Universal Robots URScript: T012_openai_gpt-oss-120b_safety_rep1.urscript

# -------------------------------------------------
# UR5e Collaborative Spot Welding Program
# Payload: 2.5 kg
# Safety: ISO 10218:2025 compliant
# -------------------------------------------------

# ---- Global Parameters ----
payload_mass = 2.5                                   # kg
payload_cog = [0,0,0]                                 # Center of gravity (m)

max_tcp_speed = 0.25                                 # m/s (250 mm/s)
max_joint_acc = 1.4                                   # rad/s^2 per joint
default_acc = 0.5                                     # m/s^2 for linear moves
default_joint_acc = 0.8                               # rad/s^2 for joint moves
default_vel = 0.2                                     # m/s (200 mm/s) default linear speed

# Workspace limits (meters) – adjust to your cell
workspace_min = [-0.8, -0.8, 0.0]                     # X, Y, Z lower bounds
workspace_max = [ 0.8,  0.8, 1.2]                     # X, Y, Z upper bounds

# ---- Safety Helper Functions ----
def check_within_workspace(p):
    # p is a pose [x, y, z, Rx, Ry, Rz]
    for i in range(3):
        if p[i] < workspace_min[i] or p[i] > workspace_max[i]:
            popup("Safety violation: Pose out of workspace bounds!", title="E-STOP", warning=True)
            halt()
    end
end

def safety_check(pose, speed):
    # Ensure speed does not exceed collaborative limit
    if speed > max_tcp_speed:
        popup("Safety violation: Speed exceeds collaborative limit!", title="E-STOP", warning=True)
        halt()
    end
    # Verify pose inside workspace
    check_within_workspace(pose)
end

def eStop_handler():
    popup("Emergency Stop triggered!", title="E-STOP", warning=True)
    halt()
end

# ---- Emergency Stop Hook ----
# URScript automatically halts on safety_stop, but we add a manual trigger for demo
def on_program_stop():
    eStop_handler()
end

# ---- Initialization ----
set_payload(payload_mass, payload_cog)                # Set payload
set_tcp(p[0,0,0,0,0,0])                               # Default TCP
set_joint_acceleration(max_joint_acc)                # Limit joint acceleration
set_joint_velocity(0.3)                               # Joint speed limit (rad/s), safe for collaborative

# ---- Define Poses ----
# Home pose (joint configuration)
home_joints = [-1.57, -1.57, 1.57, -1.57, -1.57, 0]    # rad

# Spot 1
approach_1 = p[0.300,  0.200, 0.300, 0, 3.1415, 0]    # above spot 1
weld_1    = p[0.300,  0.200, 0.100, 0, 3.1415, 0]    # descent to spot 1

# Spot 2
approach_2 = p[0.100, -0.250, 0.300, 0, 3.1415, 0]    # above spot 2
weld_2    = p[0.100, -0.250, 0.100, 0, 3.1415, 0]    # descent to spot 2

# Spot 3
approach_3 = p[-0.200, 0.150, 0.300, 0, 3.1415, 0]    # above spot 3
weld_3    = p[-0.200, 0.150, 0.100, 0, 3.1415, 0]    # descent to spot 3

# Lift pose (same X,Y as spot, safe Z)
lift_height = 0.300

# ---- Main Program ----
def main():
    # 1) Move to Home (joint move)
    safety_check(pose_from_joint(home_joints), default_vel)
    movej(home_joints, a=max_joint_acc, v=0.3)       # joint speed 0.3 rad/s (safe)

    # 2) Approach Spot 1
    safety_check(approach_1, default_vel)
    movel(approach_1, a=default_acc, v=default_vel)

    # 3) Descend to Spot 1 (welding position)
    safety_check(weld_1, 0.08)                       # 80 mm/s
    movel(weld_1, a=default_acc, v=0.08)

    # 4) Activate welding (placeholder)
    popup("Weld Spot 1 activated", title="Welding", warning=False)
    sleep(0.5)                                        # simulate weld dwell

    # 5) Lift from Spot 1
    lift_1 = pose_trans(weld_1, p[0,0,lift_height,0,0,0])
    safety_check(lift_1, 0.15)                       # 150 mm/s
    movel(lift_1, a=default_acc, v=0.15)

    # 6) Move to Spot 2
    safety_check(approach_2, default_vel)
    movel(approach_2, a=default_acc, v=default_vel)

    # 7) Descend to Spot 2
    safety_check(weld_2, 0.08)
    movel(weld_2, a=default_acc, v=0.08)

    # 8) Activate welding Spot 2
    popup("Weld Spot 2 activated", title="Welding", warning=False)
    sleep(0.5)

    # 9) Lift from Spot 2
    lift_2 = pose_trans(weld_2, p[0,0,lift_height,0,0,0])
    safety_check(lift_2, 0.15)
    movel(lift_2, a=default_acc, v=0.15)

    # 10) Move to Spot 3
    safety_check(approach_3, default_vel)
    movel(approach_3, a=default_acc, v=default_vel)

    # 11) Descend to Spot 3
    safety_check(weld_3, 0.08)
    movel(weld_3, a=default_acc, v=0.08)

    # 12) Activate welding Spot 3
    popup("Weld Spot 3 activated", title="Welding", warning=False)
    sleep(0.5)

    # 13) Lift from Spot 3
    lift_3 = pose_trans(weld_3, p[0,0,lift_height,0,0,0])
    safety_check(lift_3, 0.15)
    movel(lift_3, a=default_acc, v=0.15)

    # 14) Return Home
    safety_check(pose_from_joint(home_joints), default_vel)
    movej(home_joints, a=max_joint_acc, v=0.3)

    popup("Program completed safely.", title="Status", warning=False)
end

# ---- Helper: Convert joint vector to pose for safety_check ----
def pose_from_joint(joints):
    # Simple forward kinematics placeholder – in practice use get_forward_kin()
    # Here we assume the robot is at the pose corresponding to the joint set.
    # For safety checks we rely on workspace limits for XYZ only.
    return get_actual_pose()
end

# ---- Execute ----
main()
